(* IEC 61131-3 sources: cds-text-sync-reference-project/project-view/PLC/PLC Logic/CFC_Application/01_Object_DUT, 5 files *)

(* ---- _01_DUT_STRUCTURE.st ---- *)
TYPE _01_DUT_STRUCTURE :
STRUCT
	sName : STRING(31);        // Pump designation
	rMaxFlow : REAL := 100.0;  // Capacity limit
	xIsVFD : BOOL;            // Has Variable Frequency Drive
	diWorkingHours : DINT;    // Total service time
END_STRUCT
END_TYPE

(* ---- _01_DUT_STRUCTURE2.st ---- *)
TYPE _01_DUT_STRUCTURE2 :
STRUCT
	sName : STRING(31);        // Pump designation
	rMaxFlow : REAL := 100.0;  // Capacity limit
	xIsVFD : BOOL;            // Has Variable Frequency Drive
	diWorkingHours : DINT;    // Total service time
END_STRUCT
END_TYPE

(* ---- _02_DUT_Enumeration.st ---- *)
{attribute 'qualified_only'}
{attribute 'strict'}
TYPE _02_DUT_Enumeration :
(
	IDLE := 0,      // System waiting
	STARTING,       // Transition to running
	RUNNING,        // Active operation
	STOPPING,       // Controlled shutdown
	ERROR := 99     // Fault state
) INT;
END_TYPE

(* ---- _03_DUT_Alias.st ---- *)
TYPE _03_DUT_Alias : REAL; END_TYPE

(* ---- _04_DUT_UNION.st ---- *)
TYPE _04_DUT_UNION :
UNION
	wValue : WORD;  // Overlaps iValue
	iValue : INT;   // Overlaps wValue
END_UNION
END_TYPE
